(* IEC 61131-3 sources: trust-platform/conformance/cases/references/cfm_references_ref_to_deref_write_001, 1 file *)

(* ---- program.st ---- *)
PROGRAM Main
VAR
    target : INT := INT#5;
    ref_value : REF_TO INT := REF(target);
    observed : INT := INT#0;
    after_write : INT := INT#0;
END_VAR

observed := ref_value^;
ref_value^ := INT#8;
after_write := target;
END_PROGRAM
